RoboDK station: Simulacion2.rdk

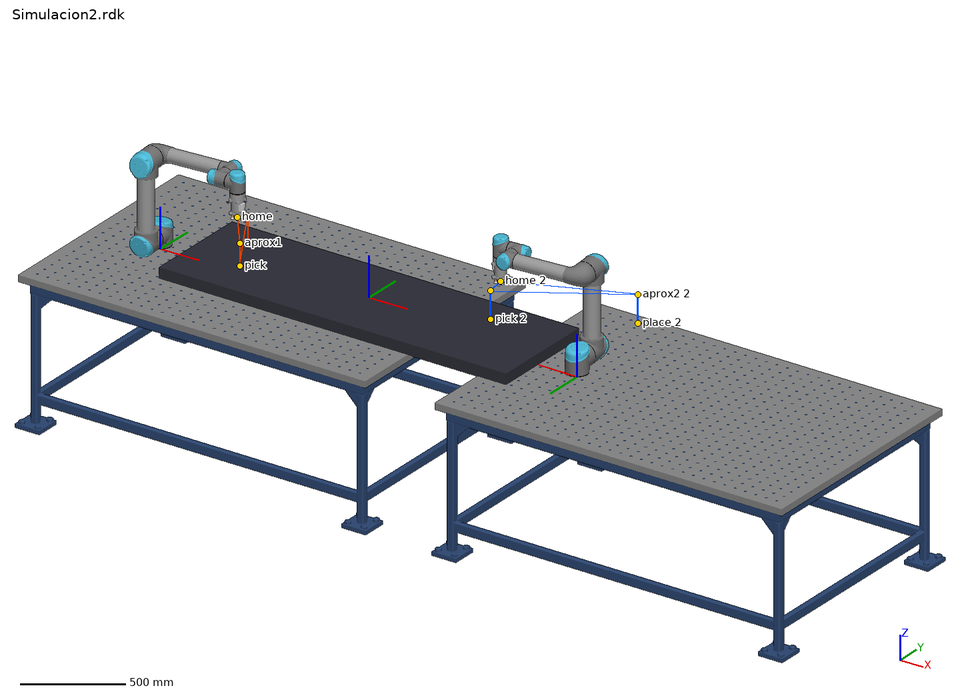
[picture v0: the station drawn from its stored meshes, robots at their saved joint values, targets as dots, program paths as lines]
Station Simulacion2 (saved by RoboDK 6.0.7). Poses are relative to the parent item; angles as X-Y-Z fixed-axis rotations.
  - frame UR5 Base at (0, -14.44, -18.09) mm
    - robot UR5: 6 axes
        modified DH rows (alpha deg, a mm, theta deg, d mm): 0, 0, 0, 89.2; 90, 0, 180, 0; 0, 425, 0, 0; 0, 392, 0, 109.3; -90, 0, 0, 94.75; 90, 0, 180, 82.5
        joint limits [-360, -360, -360, -360, -360, -360] to [360, 360, 360, 360, 360, 360]; home [0, -90, -90, 0, 90, 0]; saved at [4.15, -90, -90, -90, 90, 2.23]
      - tool SMC ZXP7A01-ZP25C-X1 Vacuum Gripper, TCP at (0, 0, 100) mm, size 70.4 x 85.4 x 102.3 mm
    - target home (Cartesian target) at (493.38, -73.79, 331.7) mm, rotated rx -180 ry 0 rz -88.08 deg; joints [4.15, -90, -90, -90, 90, 2.23] of UR5
    - target aprox1 (Cartesian target) at (508.38, -73.29, 200) mm, rotated rx -180 ry 0 rz -88.08 deg; joints [4.083, -95.038, -104.339, -70.623, 90, 2.163] of UR5
    - target pick (Cartesian target) at (508.38, -73.29, 81.7) mm, rotated rx -180 ry 0 rz -88.08 deg; joints [4.083, -103.103, -114.452, -52.445, 90, 2.163] of UR5
    - target aprox2 (Cartesian target) at (500, 0, 311.7) mm, rotated rx -180 ry 0 rz -88.08 deg; joints [51.85, -103.1, -114.45, -52.44, 90, 2.16] of UR5
    - target place (Cartesian target) at (500, 0, 161.7) mm, rotated rx -180 ry 0 rz -88.08 deg; joints [90.37, -103.09, -114.44, -52.44, 90, 2.16] of UR5
  - object Table 2000x1200x800mm at (0, 0, 0) mm, size 2020 x 1340 x 800 mm, geometry from Table-2000x1200x800mm.sld
  - Python program Crear_celda (listed below)
  - frame Conveyor Belt Base at (1200, -14.44, 61.91) mm
    - object Conveyor Belt at (0, 0, 0) mm, size 2000 x 600 x 60 mm
  - frame UR5 Base 2 at (2400, -14.44, -18.09) mm, rotated rx 0 ry 0 rz 180 deg
    - robot UR5: 6 axes
        modified DH rows (alpha deg, a mm, theta deg, d mm): 0, 0, 0, 89.2; 90, 0, 180, 0; 0, 425, 0, 0; 0, 392, 0, 109.3; -90, 0, 0, 94.75; 90, 0, 180, 82.5
        joint limits [-360, -360, -360, -360, -360, -360] to [360, 360, 360, 360, 360, 360]; home [0, -90, -90, 0, 90, 0]; saved at [4.15, -90, -90, -90, 90, 2.23]
      - tool SMC ZXP7A01-ZP25C-X1 Vacuum Gripper, TCP at (0, 0, 100) mm, size 70.4 x 85.4 x 102.3 mm
    - target home 2 (joint target) at (493.38, -73.79, 331.7) mm, rotated rx -180 ry 0 rz -88.08 deg; joints [4.15, -90, -90, -90, 90, 2.23] of UR5
    - target aprox1 2 (Cartesian target) at (500, 0, 311.7) mm, rotated rx 180 ry 0 rz -88.08 deg; joints [12.627, -90.225, -92.699, -87.076, 90, 10.707] of UR5
    - target pick 2 (Cartesian target) at (500, 0, 161.7) mm, rotated rx 180 ry 0 rz -88.08 deg; joints [12.627, -95.276, -110.134, -64.591, 90, 10.707] of UR5
    - target aprox2 2 (Cartesian target) at (0, -500, 231.7) mm, rotated rx 180 ry 0 rz -88.08 deg; joints [-77.373, -91.897, -102.848, -75.256, 90, -79.293] of UR5
    - target place 2 (Cartesian target) at (0, -500, 81.7) mm, rotated rx 180 ry 0 rz -88.08 deg; joints [77.373, 23.12, -83.828, -209.292, 90, 75.453] of UR5
  - object Table 2 at (2400, 0, 0) mm, size 2020 x 1340 x 800 mm, geometry from Table-2000x1200x800mm.sld
  - program Prog2 (10 instructions, listed below)
  - program Prog1 (8 instructions, listed below)
  - object Box 24x16in (Closed) at (2400, 485.56, -86.39) mm, rotated rx 0 ry 0 rz -88.08 deg, size 99.5 x 152.5 x 66.9 mm, geometry from Box-24x16in-Closed.sld
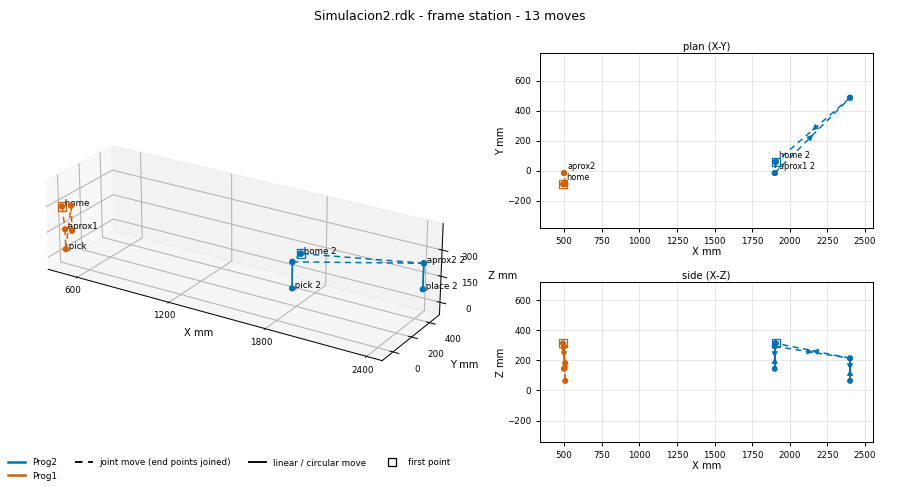
[picture p0: tool path of Simulacion2.rdk in frame station, 13 of 13 moves have a stored position in this frame; points joined in program order, loops and branches not executed]

--- Python program Crear_celda ---
from robodk.robolink import *
from robodk.robomath import *
import ast

GAP = 2400
BELT_START = 500
BELT_END = 1900
CONV_DX = 1200
CONV_DY = 0
CONV_ROT_Z = 0
CONV_Z_OFF = 80
PLACE2_DX = 0
PLACE2_DY = 500
APPROACH = 150
BOX_H = 150
STEPS = 100

RDK = Robolink()
station = RDK.ActiveStation()

def buscar(tipo, empieza=None, contiene=None, excluir=()): return next((it for it in RDK.ItemList(tipo) if it.Name() not in excluir and ((empieza and it.Name().startswith(empieza)) or (contiene and contiene.lower() in it.Name().lower()))), None)
def hijos(item, tipo): return [c for c in item.Childs() if c.Type() == tipo]

base1 = RDK.Item('UR5 Base', ITEM_TYPE_FRAME)
robot1 = hijos(base1, ITEM_TYPE_ROBOT)[0]
tool1 = hijos(robot1, ITEM_TYPE_TOOL)[0]
tg = {c.Name(): c for c in hijos(base1, ITEM_TYPE_TARGET)}
home1, aprox1, pick1, aprox2, place1 = [tg[n] for n in ('home', 'aprox1', 'pick', 'aprox2', 'place')]

table1 = buscar(ITEM_TYPE_OBJECT, empieza='Table', excluir=('Table 2',))
box = buscar(ITEM_TYPE_OBJECT, empieza='Box')
conv = buscar(ITEM_TYPE_FRAME, contiene='conveyor')
if table1 is None or box is None or conv is None: raise Exception('No encuentro la mesa (Table...), la caja (Box...) o la banda (Conveyor...).')

in_tool = box.Parent().Type() == ITEM_TYPE_TOOL
tcp_now = robot1.PoseAbs() * robot1.SolveFK(robot1.Joints()) * tool1.PoseTool()
T = invH(tcp_now) * box.PoseAbs() if in_tool else None
if in_tool: RDK.setParam('T_TCP_BOX', repr(T.tolist())); box.setParentStatic(station)
saved = RDK.getParam('T_TCP_BOX')
if not in_tool: T = Mat(ast.literal_eval(saved)) if saved else transl(0, 0, BOX_H) * rotx(pi)

base2 = RDK.Item('UR5 Base 2', ITEM_TYPE_FRAME)
nombres = {'home': 'home 2', 'aprox1': 'aprox1 2', 'pick': 'pick 2', 'aprox2': 'aprox2 2', 'place': 'place 2'}
if not base2.Valid(): base1.Copy(); base2 = RDK.Paste(); base2.setName('UR5 Base 2'); [ch.setName(nombres[ch.Name()]) for ch in base2.Childs() if ch.Name() in nombres]; table1.Copy(); RDK.Paste().setName('Table 2')

table2 = RDK.Item('Table 2', ITEM_TYPE_OBJECT)
robot2 = hijos(base2, ITEM_TYPE_ROBOT)[0]
tool2 = hijos(robot2, ITEM_TYPE_TOOL)[0]
t2 = {c.Name(): c for c in hijos(base2, ITEM_TYPE_TARGET)}
home2, aprox12, pick2, aprox22, place2 = [t2[n] for n in ('home 2', 'aprox1 2', 'pick 2', 'aprox2 2', 'place 2')]

B1 = base1.PoseAbs()
p1 = B1.Pos()
surf_z = p1[2]
base2.setPoseAbs(transl(GAP, 0, 0) * B1 * rotz(pi))
table2.setPoseAbs(transl(GAP, 0, 0) * table1.PoseAbs())
conv.setPoseAbs(transl(p1[0] + CONV_DX, p1[1] + CONV_DY, surf_z + CONV_Z_OFF) * rotz(CONV_ROT_Z * pi / 180))

B0 = pick1.PoseAbs() * T
box.setPoseAbs(B0)
dz = B0.Pos()[2] - surf_z
R0 = invH(transl(*B0.Pos())) * B0
zb = surf_z + dz + CONV_Z_OFF
B_start = transl(p1[0] + BELT_START, p1[1], zb) * R0
B_end = transl(p1[0] + BELT_END, p1[1], zb) * R0
B_dest = transl(p1[0] + GAP + PLACE2_DX, p1[1] + PLACE2_DY, surf_z + dz) * R0

place1_tcp = B_start * invH(T)
place1.setPoseAbs(place1_tcp)
aprox2.setPoseAbs(transl(0, 0, APPROACH) * place1_tcp)

T2 = invH(rotz(pi)) * T
pick2_tcp = B_end * invH(T) * rotz(pi)
place2_tcp = B_dest * invH(T2)
for t, pose in ((pick2, pick2_tcp), (place2, place2_tcp), (aprox12, transl(0, 0, APPROACH) * pick2_tcp), (aprox22, transl(0, 0, APPROACH) * place2_tcp)): t.setAsCartesianTarget(); t.setPoseAbs(pose)
home2.setAsJointTarget()
home2.setJoints(home1.Joints())

if not RDK.Item('Prog2', ITEM_TYPE_PROGRAM).Valid(): prog2 = RDK.AddProgram('Prog2', robot2); prog2.setPoseFrame(base2); prog2.setPoseTool(tool2); prog2.MoveJ(home2); prog2.MoveJ(aprox12); prog2.MoveL(pick2); prog2.MoveL(aprox12); prog2.MoveJ(aprox22); prog2.MoveL(place2); prog2.MoveL(aprox22); prog2.MoveJ(home2)

robot1.setPoseFrame(base1)
robot1.setPoseTool(tool1)
robot2.setPoseFrame(base2)
robot2.setPoseTool(tool2)

robot1.MoveJ(home1)
robot1.MoveJ(aprox1)
robot1.MoveL(pick1)
box.setParentStatic(tool1)
robot1.MoveL(aprox1)
robot1.MoveJ(aprox2)
robot1.MoveL(place1)
box.setParentStatic(station)
robot1.MoveL(aprox2)
robot1.MoveJ(home1)

for i in range(STEPS + 1): box.setPoseAbs(transl(p1[0] + BELT_START + (BELT_END - BELT_START) * i / STEPS, p1[1], zb) * R0); RDK.Render(True); pause(0.02)

robot2.MoveJ(home2)
robot2.MoveJ(aprox12)
robot2.MoveL(pick2)
box.setParentStatic(tool2)
robot2.MoveL(aprox12)
robot2.MoveJ(aprox22)
robot2.MoveL(place2)
box.setParentStatic(station)
robot2.MoveL(aprox22)
robot2.MoveJ(home2)
print('Listo.')

--- program Prog2 (robot UR5) ---
  Est. Ref.: UR5 Base 2
  Est. herr: SMC ZXP7A01-ZP25C-X1 Vacuum Gripper
  MoveJ (home 2)
  MoveJ (aprox1 2)
  MoveL (pick 2)
  MoveL (aprox1 2)
  MoveJ (aprox2 2)
  MoveL (place 2)
  MoveL (aprox2 2)
  MoveJ (home 2)

--- program Prog1 (robot UR5) ---
  Est. Ref.: UR5 Base
  Est. herr: SMC ZXP7A01-ZP25C-X1 Vacuum Gripper
  MoveJ (home)
  MoveJ (aprox1)
  MoveJ (pick)
  Adjuntar a SMC ZXP7A01-ZP25C-X1 Vacuum Gripper
  MoveJ (aprox2)
  MoveJ (place)
